(*
SPDX-FileCopyrightText: © 2026 Oleksandr Tiutyk <trofimich@gmail.com>
SPDX-License-Identifier: MIT
License: https://opensource.org/license/mit
*)

(*!
<summary>Names preparation and write-failure checks for a file opened for reading.</summary>
<description>
Steps belong to one test scenario; values are not a serialized protocol. The first member is the initial
preparation step. Test completion and failure cleanup are tracked separately.
</description>
*)
{attribute 'qualified_only'}
{attribute 'strict'}
{attribute 'to_string'}
TYPE READ_ONLY_FILE_TEST_STEP :
(
	CREATE_FILE,
	OPEN_FILE_FOR_READING,
	CHECK_WRITE_FAILURE
);
END_TYPE

(* stored: Version 1.1.0.1
   DUT READ_ONLY_FILE_TEST_STEP: Id {efd85a05-418b-4ead-8fd7-a88688323289} *)
